TYPE ST_PersistentInner :
STRUCT
	nCount : INT;
	fOffset : LREAL;
END_STRUCT
END_TYPE

(* stored: Version 1.1.0.1
   DUT ST_PersistentInner: Id {3f6a1c52-8d7e-4b0a-9a41-5c2e7d9b1a01} *)
